Fanuc KAREL source: KA00129.KL

PROGRAM KA00129
%NOLOCKGROUP
VAR
  SRC: ARRAY[2] OF BYTE
  DST: VECTOR
BEGIN
  SRC[1] = 2
  DST = SRC[1]
END KA00129
